INTERFACE I_Light EXTENDS I_Device

PROPERTY IsOn : BOOL
GET
END_GET
END_PROPERTY

METHOD TurnOn
END_METHOD

METHOD TurnOff
END_METHOD

METHOD Toggle
END_METHOD

METHOD SetBrightness
VAR_INPUT
    nBrightness : UINT;
END_VAR
END_METHOD

END_INTERFACE

(* stored: Version 1.1.0.1
   Itf I_Light: Id {A1A1A1A1-A1A1-41A1-81A1-A1A1A1A1A1A0}
   Property IsOn: Id {A1A1A1A1-A1A1-41A1-81A1-A1A1A1A1A1A1}
   Get Get: Id {A1A1A1A1-A1A1-41A1-81A1-A1A1A1A1A1A2}
   Method TurnOn: Id {A1A1A1A1-A1A1-41A1-81A1-A1A1A1A1A1A3}
   Method TurnOff: Id {A1A1A1A1-A1A1-41A1-81A1-A1A1A1A1A1A4}
   Method Toggle: Id {A1A1A1A1-A1A1-41A1-81A1-A1A1A1A1A1A5}
   Method SetBrightness: Id {A1A1A1A1-A1A1-41A1-81A1-A1A1A1A1A1A6} *)
